Staubli VAL3: send.pgx

program send()
  local num i
  local bool l_bEnabling
  local bool l_bErr
  local bool l_bLastPower
  local bool l_bMcpEstop
  local num l_i
begin
  //远程模式
  dOutWorkingMode=rs:bIsRemoteAuto
  //上电
  dOutIsPowerd=isPowered()
  //程序运行
  dOutCycle=rs:bIsCycle
  //机器人报警
  dOutError=rs:bIsError
  //机器人急停
  dOutEstop=rs:bIsEstop
  //机器人在原点
  dOutIsHome=rs:bIsHome
  //机器人通讯故障
  if ioStatus(dOutIsHome)<0
    rs:bIsError=true
  endIf
end
